// TIA Portal V20 export
Screen "OP04Pop-up_PRBWork"  274x160
  ScreenItem "Text field TG Status" at 3,5 size 273x47  Type=HmiTextBox
  ScreenItem "Cancel Mode" at 197,8 size 76x42  Type=HmiButton
  ScreenItem "Rectangle TG1" at 6,57 size 265x29  Type=HmiRectangle
  ScreenItem "Textfeld_1" at 11,62 size 21x20  Type=HmiTextBox
  ScreenItem "Textfeld_2" at 52,61 size 245x20  Type=HmiTextBox
  ScreenItem "Rectangle TG1_1" at 6,89 size 265x29  Type=HmiRectangle
  ScreenItem "Textfeld_5" at 11,93 size 21x20  Type=HmiTextBox
  ScreenItem "Rectangle TG1_5" at 6,122 size 265x29  Type=HmiRectangle
  ScreenItem "Textfeld_3" at 52,93 size 245x20  Type=HmiTextBox
  ScreenItem "Textfeld_11" at 52,125 size 275x20  Type=HmiTextBox
  ScreenItem "Textfeld_16" at 11,129 size 21x20  Type=HmiTextBox
  ScreenItem "Line_1" at 39,55 size 1x101  Type=HmiLine
